FUNCTION_BLOCK SortingHomeConditions (* Sorting-only architecture following Distribution and tutorial modules 1-4 *)
  (* Standard: 61499-2 *)
  (* Version 2.0, 2026-11-09, sorting2n, sorting2n *)
  PACKAGE Main;
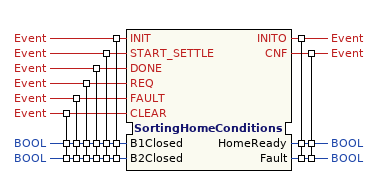
  EVENT_INPUT
    INIT WITH B1Closed, B2Closed;
    START_SETTLE WITH B1Closed, B2Closed;
    DONE WITH B1Closed, B2Closed;
    REQ WITH B1Closed, B2Closed;
    FAULT WITH B1Closed, B2Closed;
    CLEAR WITH B1Closed, B2Closed;
  END_EVENT
  EVENT_OUTPUT
    INITO WITH HomeReady, Fault;
    CNF WITH HomeReady, Fault;
  END_EVENT
  VAR_INPUT
    B1Closed : BOOL;
    B2Closed : BOOL;
  END_VAR
  VAR_OUTPUT
    HomeReady : BOOL;
    Fault : BOOL;
  END_VAR
  VAR
    Elapsed : BOOL;
  END_VAR
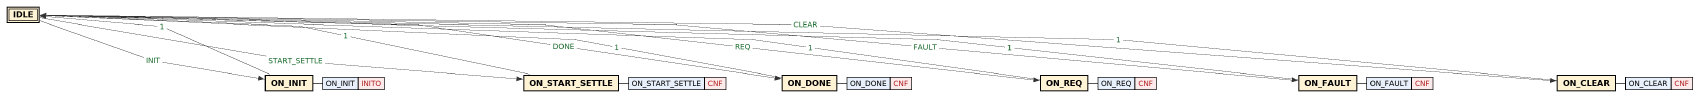
  EC_STATES
    IDLE;
    ON_INIT : ON_INIT -> INITO;
    ON_START_SETTLE : ON_START_SETTLE -> CNF;
    ON_DONE : ON_DONE -> CNF;
    ON_REQ : ON_REQ -> CNF;
    ON_FAULT : ON_FAULT -> CNF;
    ON_CLEAR : ON_CLEAR -> CNF;
  END_STATES
  EC_TRANSITIONS
    IDLE TO ON_INIT := INIT;
    ON_INIT TO IDLE := 1;
    IDLE TO ON_START_SETTLE := START_SETTLE;
    ON_START_SETTLE TO IDLE := 1;
    IDLE TO ON_DONE := DONE;
    ON_DONE TO IDLE := 1;
    IDLE TO ON_REQ := REQ;
    ON_REQ TO IDLE := 1;
    IDLE TO ON_FAULT := FAULT;
    ON_FAULT TO IDLE := 1;
    IDLE TO ON_CLEAR := CLEAR;
    ON_CLEAR TO IDLE := 1;
  END_TRANSITIONS
  ALGORITHM ON_INIT IN ST:
Elapsed := FALSE; HomeReady := FALSE; Fault := FALSE;
  END_ALGORITHM
  ALGORITHM ON_START_SETTLE IN ST:
Elapsed := FALSE; HomeReady := FALSE;
  END_ALGORITHM
  ALGORITHM ON_DONE IN ST:
Elapsed := TRUE; HomeReady := B1Closed AND B2Closed;
  END_ALGORITHM
  ALGORITHM ON_REQ IN ST:
HomeReady := Elapsed AND B1Closed AND B2Closed AND NOT Fault;
  END_ALGORITHM
  ALGORITHM ON_FAULT IN ST:
Fault := TRUE; HomeReady := FALSE;
  END_ALGORITHM
  ALGORITHM ON_CLEAR IN ST:
Fault := FALSE; Elapsed := FALSE; HomeReady := FALSE;
  END_ALGORITHM
END_FUNCTION_BLOCK
